(* IEC 61131-3 sources: 2026_Projet_YGO_ExcavatriceDragage/CODE_BACKUP/CODE_20260902_JoyAvantHoming_v0.6.27/I_TRANSLATION/_TYPES, 5 files *)

(* ---- E_TranslationFinalInterlockReason.st ---- *)
(* =======================================================================
   🛡️ E_TranslationFinalInterlockReason — Raisons d'interlock M3
   ───────────────────────────────────────────────────────────────
   🎯 Rôle : Énumération des raisons de blocage de la barrière finale M3
   📄 Doc métier : DOC/AF/AF_Partie-11_Fonction_Translation_v2.3.md
   ======================================================================= *)
{attribute 'qualified_only'}
TYPE E_TranslationFinalInterlockReason :
(
    NONE := 0,
    BRAKE_COMMAND_NOT_CONFIRMED := 1,
    RESTART_INHIBITED := 2
);
END_TYPE

(* ---- ST_fbTranslation_Cfg.st ---- *)
(* ═══════════════════════════════════════════════════════════════
   ⚙️ ST_fbTranslation_Cfg — Configuration regroupée de FB_Translation
   ───────────────────────────────────────────────────────────────
   📐 NC-110 / G380 : pattern « Cfg : ST_fb<Fb>_Cfg » (comme FB_Winch
      avec Config : ST_fbWinch_Cfg). Regroupe en UN point d'interface les
      ~13 scalaires `[CFG]` qui étaient des VAR_INPUT plates de FB_Translation.
   🎯 Un seul sourcing : PRG_05_Translation assemble ce struct depuis la
      source unique GVL_PERSISTENT (§ source propre documentée ci-dessous).
   📤 Producteur : PRG_05_Translation (câblage).
   📥 Consommateur : FB_Translation (Cfg, lecture seule).
   📄 Doc : DOC/AF/AF_Partie-11_Fonction_Translation_v2.3.md
   ═══════════════════════════════════════════════════════════════ *)

TYPE ST_fbTranslation_Cfg :
STRUCT
    // === RAMPES VITESSE (%/s) ===
    CfgRampAccelRate            : REAL := 20.0;   // --> [CFG] Accélération
    CfgRampDecelNormalRate      : REAL := 40.0;   // --> [CFG] Décélération normale
    CfgRampDecelFastRate        : REAL := 100.0;  // --> [CFG] Décélération RAPIDE (SafeStop)
    DirectionInterlockDelay     : TIME := T#200ms; // --> [CFG] Délai avant changement de sens à l'arrêt

    // === VITESSES RÉDUITES D'APPROCHE (Hz) ===
    ApproachSpeedTremieHz       : REAL := 10.0;   // --> [CFG] Approche Trémie (Direction=1)
    ApproachSpeedMaintenanceHz  : REAL := 10.0;   // --> [CFG] Approche Maintenance (Direction=-1)
    ApproachSpeedP1Hz           : REAL := 10.0;   // --> [CFG] Approche P1 (Direction=-1)

    // === ÉCHELLE VARIATEUR ===
    DriveFreqScaleMaxHz         : REAL := 60.0;   // --> [CFG] Échelle 0..100 % → MaxHz

    // === COMMUN / FREIN ===
    CaptorDebounce              : TIME := T#100ms; // --> [CFG] Filtrage capteur position cible
    BrakeDelayContactClose      : TIME := T#100ms; // --> [CFG] Voir FB_Brake
    BrakeDelayMagnetise         : TIME := T#100ms; // --> [CFG] Voir FB_Brake
    BrakeDelayMotorDecel        : TIME := T#500ms; // --> [CFG] Voir FB_Brake
    BrakeFeedbackTimeout        : TIME := T#300ms; // --> [CFG] Strictement sous watchdog final 500 ms
END_STRUCT
END_TYPE

(* ---- ST_fbTranslationCmdArbitration_Cfg.st ---- *)
(* ═══════════════════════════════════════════════════════════════
   ⚙️ ST_fbTranslationCmdArbitration_Cfg — Config translation M3
   ───────────────────────────────────────────────────────────────
   🎯 Rôle : Config statique de FB_TranslationCmdArbitrationM3.
       Porte la fréquence max (échelle FreqPct) — paramètre de config,
       pas un fait de gating (I5). Le Context ne garde que les faits
       de gating (HeightInterlockOk).
   📤 Producteur : PRG_05_Translation (câblage).
   📄 Doc : DOC/AF/AF_Partie-11_Fonction_Translation_v2.3.md
   🔌 Source : GVL_PERSISTENT._TranslationMaxFreq_Hz (source unique).
   ═══════════════════════════════════════════════════════════════ *)

TYPE ST_fbTranslationCmdArbitration_Cfg :
STRUCT
    MaxFreq_Hz : REAL;  // --> [CFG] Fréquence max (échelle FreqPct, _TranslationMaxFreq_Hz)
END_STRUCT
END_TYPE

(* ---- ST_fbTranslationCmdArbitration_Context.st ---- *)
(* ═══════════════════════════════════════════════════════════════
   🧩 ST_fbTranslationCmdArbitration_Context — Contexte de gating M3
   ───────────────────────────────────────────────────────────────
   🎯 Rôle : Encapsuler les faits de gating consommés par FB_TranslationCommandArbitration
       (interlock hauteur M1/M2).
       La fréquence max (config) vit dans ST_fbTranslationCmdArbitration_Cfg (I5).
   📤 Producteur : PRG_05_Translation (câblage).
   📄 Doc : DOC/AF/AF_Partie-11_Fonction_Translation_v2.3.md
   ═══════════════════════════════════════════════════════════════ *)

TYPE ST_fbTranslationCmdArbitration_Context :
STRUCT
    HeightInterlockOk : BOOL;  // --> [SAFE] Hauteur mini M1/M2 OK (anti-collision translation)
END_STRUCT
END_TYPE

(* ---- ST_fbTranslationCmdArbitration_IHM.st ---- *)
(* ═══════════════════════════════════════════════════════════════
   🎛️ ST_fbTranslationCmdArbitration_IHM — Entrées IHM de l'arbitrage M3
   ───────────────────────────────────────────────────────────────
   🎯 Rôle : Encapsuler les commandes IHM consommées par FB_TranslationCommandArbitration
       (boutons, sélecteur positionnement, consigne fréquence).
       Le toggle joystick maître global (Modes.Cmd.TglJoystickMaster) est passé en
       paramètre séparé du FB (I4 — factorisation, source unique GVL_IHM.Modes.Cmd).
   📤 Producteur : PRG_05_Translation (câblage GVL_IHM).
   📄 Doc : DOC/AF/AF_Partie-11_Fonction_Translation_v2.3.md
   ═══════════════════════════════════════════════════════════════ *)

TYPE ST_fbTranslationCmdArbitration_IHM :
STRUCT
    BtnTremie         : BOOL;  // --> [CMD] Bouton translation vers Trémie (TranslationM3.Cmd.BtnTremie, ex-BtnFwd)
    BtnMaintenance    : BOOL;  // --> [CMD] Bouton translation vers Maintenance (TranslationM3.Cmd.BtnMaintenance, ex-BtnRev)
    SelPositioning    : BOOL;  // --> [CMD] Sélecteur positionnement (TranslationM3.Cmd.SelPositioning)
    SetFreq_Hz        : REAL;  // --> [CMD] Consigne fréquence (TranslationM3.Cmd.SetFreq_Hz)
    BypassGlobal      : BOOL;  // --> [TST] Bypass global translation (TranslationM3.Bypass.Global)
END_STRUCT
END_TYPE
